Fanuc KAREL source: KA00202.KL

PROGRAM KA00202
%NOLOCKGROUP
VAR
  SRC: ARRAY[4] OF VECTOR
  DST: ARRAY[4] OF STRING[20]
BEGIN
  DST = SRC
END KA00202
